ADAPTER EventAdapter (* Adapter with event and data interfaces *)
  (* Standard: 61499-1; Description: Copyright (c) 2026 Martin Erich Jobst This program and the accompanying materials are made available under the terms of the Eclipse Public License 2.0 which is available at https://www.eclipse.org/legal/epl-2.0/ SPDX-License-Identifier: EPL-2.0 *)
  (* Version 1.0, 2026-10-23, Martin Jobst *)
  {SET_ATTRIBUTE(IntegerAttribute, 4)}
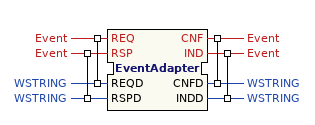
  EVENT_INPUT
    REQ WITH REQD;
    RSP WITH RSPD;
  END_EVENT
  EVENT_OUTPUT
    CNF WITH CNFD;
    IND WITH INDD;
  END_EVENT
  VAR_INPUT
    REQD : WSTRING; (* Request data *)
    RSPD : WSTRING; (* Response data *)
  END_VAR
  VAR_OUTPUT
    CNFD : WSTRING; (* Confirmation data *)
    INDD : WSTRING; (* Indication data *)
  END_VAR
  SERVICE PLUG/SOCKET (* Adapter with only events *)
    SEQUENCE request_confirm
      SOCKET.REQ(REQD) -> PLUG.REQ(REQD);
      PLUG.CNF(CNFD) -> SOCKET.CNF(CNFD);
    END_SEQUENCE
    SEQUENCE indication_response
      PLUG.IND(INDD) -> SOCKET.IND(INDD);
      SOCKET.RSP(RSPD) -> PLUG.RSP(RSPD);
    END_SEQUENCE
  END_SERVICE
END_ADAPTER
